// Base of the HalfBROTTests suites: Check() is a TcUnit assertion that also notes a failed check in GVL_Diag.sFailures
// (printed by tools/Run-Tests.ps1, TcUnit itself writes the failure text only to the ADS log). The test method sets
// sCurrent to its name first.
FUNCTION_BLOCK FB_TestBase EXTENDS TcUnit.FB_TestSuite
VAR
	sCurrent	: STRING(80);
END_VAR

METHOD Check
VAR_INPUT
	bCondition	: BOOL;
	sMessage	: STRING(255);
END_VAR
AssertTrue(Condition := bCondition, Message := sMessage);
F_Note(bFailed := NOT bCondition, sText := CONCAT(sCurrent, sMessage));
END_METHOD

END_FUNCTION_BLOCK

(* stored: Version 1.1.0.1, ProductVersion 3.1.4024.15
   POU FB_TestBase: Id {beb16b7e-96a2-53a3-a263-4d8829c174ef}, SpecialFunc None
   Method Check: Id {eb2f27e5-d226-5090-a92c-4481eb08b27d} *)
